  rq_init_comm_if_connected(9, "1")
  rq_init_comm_if_connected(2, "2")
  rq_init_comm_if_connected(3, "3")
  rq_init_comm_if_connected(4, "4")
  rq_print_connected_grippers()
  rq_gripper_communication_thread = run rq_gripper_communication()
  set_closed_norm(97.6470588235294, "1")
  set_open_norm(1.1764705882352942, "1")
  set_closed_mm(0.0, "1")
  set_open_mm(53.0, "1")
  set_closed_norm(100.0, "2")
  set_open_norm(0.0, "2")
  set_closed_mm(0.0, "2")
  set_open_mm(50.0, "2")
  set_closed_norm(100.0, "3")
  set_open_norm(0.0, "3")
  set_closed_mm(0.0, "3")
  set_open_mm(50.0, "3")
  set_closed_norm(100.0, "4")
  set_open_norm(0.0, "4")
  set_closed_mm(0.0, "4")
  set_open_mm(50.0, "4")
  rq_current_limit_enabled = False
  while(not rq_gripper_communication_thread_started):
      sleep(0.008)
  end
  # end: URCap Installation Node
  step_count_652fcfe5_f3e5_4323_a28e_c4dd7c99f65c = 0.0
  thread Step_Counter_Thread_2d5c0d0e_2884_4a5b_ab92_48b0595c18f1():
    while (True):
      step_count_652fcfe5_f3e5_4323_a28e_c4dd7c99f65c = step_count_652fcfe5_f3e5_4323_a28e_c4dd7c99f65c + 1.0
      sync()
    end
  end
  run Step_Counter_Thread_2d5c0d0e_2884_4a5b_ab92_48b0595c18f1()
  global DEV_CEN_PosRtr=0
  $ 2 "BeforeStart"
  $ 3 "Centrifuge≔rpc_factory('xmlrpc','http://192.168.12.125:50002')"
  global Centrifuge=rpc_factory("xmlrpc","http://192.168.12.125:50002")
  $ 4 "Action≔'What to do?'"
  global Action=request_integer_from_primary_client("What to do?")
  $ 5 "Robot Program"
  $ 6 "Handling"
  $ 44 "'===================='"
  # '===================='
  $ 45 "Switch Action"
  switch_1 = Action
  $ 46 "Case 5"
  if (5 == switch_1):
    $ 47 "Open"
    $ 48 "Centrifuge.open_hatch()"
    Centrifuge.open_hatch()
  elif (6 == switch_1):
    $ 49 "Case 6"
    $ 50 "Close"
    $ 51 "Centrifuge.close_hatch()"
    Centrifuge.close_hatch()
  elif (7 == switch_1):
    $ 52 "Case 7"
    $ 53 "Load"
    $ 54 "DEV_CEN_CmdRslt≔Centrifuge.move_rotor(DEV_CEN_PosRtr)"
    global DEV_CEN_CmdRslt=Centrifuge.move_rotor(DEV_CEN_PosRtr)
    $ 55 "If JNT_S≠[0,0,0,0,0,0]"
    if (JNT_S != [0,0,0,0,0,0]):
      $ 56 "MoveJ"
      $ 57 "JNT_S" "breakAfter"
      movej(JNT_S, a=1.3962634015954636, v=1.5707963267948966, r=0.05)
    end
    $ 58 "MoveJ"
    $ 59 "If PSE_A_H≠p[0,0,0,0,0,0]"
    if (PSE_A_H != p[0,0,0,0,0,0]):
      $ 60 "PSE_A_H" "breakAfter"
      movej(pose_trans(FRM_Reference, PSE_A_H), a=1.3962634015954636, v=1.5707963267948966, r=0.02)
    end
    $ 61 "PSE_A" "breakAfter"
    movej(pose_trans(FRM_Reference, PSE_A), a=1.3962634015954636, v=1.5707963267948966)
    $ 62 "If Centrifuge.posreached(DEV_CEN_PosRtr)"
    if (Centrifuge.posreached(DEV_CEN_PosRtr)):
      $ 63 "MoveL"
      $ 64 "If PSE_T_H≠p[0,0,0,0,0,0]"
      if (PSE_T_H != p[0,0,0,0,0,0]):
        $ 65 "PSE_T_H" "breakAfter"
        movel(pose_trans(FRM_Reference, PSE_T_H), a=1.2, v=0.3)
      end
      $ 66 "PSE_T" "breakAfter"
      global move_thread_flag_66=0
      thread move_thread_66():
        enter_critical
        move_thread_flag_66 = 1
        movel(pose_trans(FRM_Reference, PSE_T), a=1.2, v=0.075)
        move_thread_flag_66 = 2
        exit_critical
      end
      move_thread_flag_66 = 0
      move_thread_han_66 = run move_thread_66()
      while (True):
        local targetTcpDirection=get_target_tcp_speed()
        local stepsToRetract=tool_contact(direction=targetTcpDirection)
        if (stepsToRetract > 0):
          kill move_thread_han_66
          stopl(0.5)
          local backTrackMovement=get_actual_joint_positions_history(stepsToRetract)
          local contactPose=get_forward_kin(backTrackMovement)
          local posDir=[targetTcpDirection[0],targetTcpDirection[1],targetTcpDirection[2]]
          local retractTo=contactPose
          if (norm(posDir) > 1e-6):
            local normalizedPosDir=normalize(posDir)
            local additionalRetraction=p[normalizedPosDir[0] * 0.001, normalizedPosDir[1] * 0.001, normalizedPosDir[2] * 0.001, 0, 0, 0]
            retractTo = pose_sub(contactPose, additionalRetraction)
          end
          movel(retractTo, a=0.5, v=0.1)
          $ 67 "Until (tool_contact_detection)"
          $ 68 "EOAT"
          # begin: URCap Program Node
          #   Source: Robotiq_Grippers, 3.11.2.92906, Robotiq Inc.
          #   Type: Gripper
          $ 69 "Gripper Move5mm (1)"
          if not(gripper_connected[0]):
            popup("Gripper 1 must be connected to run this program.", "No connection", False, True, True)
          end
          if not(rq_is_gripper_activated("1")):
            popup("Gripper 1 is not activated. Go to Installation tab > Gripper to activate it and run the program again.", "Not activated", False, True, True)
          end
          rq_set_pos_spd_for(226, 128, 64, "1")
          rq_wait_pos_spe_for_request(226, 128, 64, "1")
          rq_go_to("1")
          rq_wait("1")
          # end: URCap Program Node
          $ 70 "Force"
          sleep(0.02)
          zero_ftsensor()
          force_mode(tool_pose(), [0, 0, 0, 0, 0, 1], [0.0, 0.0, 0.0, 0.0, 0.0, 0.0], 2, [0.1, 0.1, 0.1, 0.3490658503988659, 0.3490658503988659, 3.141592653589793])
          $ 71 "PSE_T" "noBreak"
          movel(pose_trans(FRM_Reference, PSE_T), a=1.2, v=0.01)
          end_force_mode()
          stopl(5.0)
          break
        end
        sleep(1.0E-10)
        if (move_thread_flag_66 > 1):
          join move_thread_han_66
          break
        end
        sync()
      end
      $ 72 "EOAT"
      # begin: URCap Program Node
      #   Source: Robotiq_Grippers, 3.11.2.92906, Robotiq Inc.
      #   Type: Gripper
      $ 73 "Gripper Move15mm (1)"
      if not(gripper_connected[0]):
        popup("Gripper 1 must be connected to run this program.", "No connection", False, True, True)
      end
      if not(rq_is_gripper_activated("1")):
        popup("Gripper 1 is not activated. Go to Installation tab > Gripper to activate it and run the program again.", "Not activated", False, True, True)
      end
      rq_set_pos_spd_for(179, 128, 128, "1")
      rq_wait_pos_spe_for_request(179, 128, 128, "1")
      rq_go_to("1")
      rq_wait("1")
      # end: URCap Program Node
      $ 74 "If PSE_R_H≠p[0,0,0,0,0,0]"
      if (PSE_R_H != p[0,0,0,0,0,0]):
        $ 75 "PSE_R" "breakAfter"
        movel(pose_trans(FRM_Reference, PSE_R), a=1.2, v=0.3, r=0.01)
        $ 76 "PSE_R_H" "breakAfter"
        movel(pose_trans(FRM_Reference, PSE_R_H), a=1.2, v=0.3)
      else:
        $ 77 "Else" "noBreak"
        $ 78 "PSE_R" "breakAfter"
        movel(pose_trans(FRM_Reference, PSE_R), a=1.2, v=0.3)
      end
    end
  elif (8 == switch_1):
    $ 79 "Case 8"
    $ 80 "Unload"
    $ 81 "DEV_CEN_CmdRslt≔Centrifuge.move_rotor(DEV_CEN_PosRtr)"
    global DEV_CEN_CmdRslt=Centrifuge.move_rotor(DEV_CEN_PosRtr)
    $ 82 "If JNT_S≠[0,0,0,0,0,0]"
    if (JNT_S != [0,0,0,0,0,0]):
      $ 83 "MoveJ"
      $ 84 "JNT_S" "breakAfter"
      movej(JNT_S, a=1.3962634015954636, v=1.5707963267948966, r=0.05)
    end
    $ 85 "MoveJ"
    $ 86 "If PSE_A_H≠p[0,0,0,0,0,0]"
    if (PSE_A_H != p[0,0,0,0,0,0]):
      $ 87 "PSE_A_H" "breakAfter"
      movej(pose_trans(FRM_Reference, PSE_A_H), a=1.3962634015954636, v=1.5707963267948966, r=0.02)
    end
    $ 88 "PSE_A" "breakAfter"
    movej(pose_trans(FRM_Reference, PSE_A), a=1.3962634015954636, v=1.5707963267948966)
    $ 89 "EOAT"
    # begin: URCap Program Node
    #   Source: Robotiq_Grippers, 3.11.2.92906, Robotiq Inc.
    #   Type: Gripper
    $ 90 "Gripper Move15mm (1)"
    if not(gripper_connected[0]):
      popup("Gripper 1 must be connected to run this program.", "No connection", False, True, True)
    end
    if not(rq_is_gripper_activated("1")):
      popup("Gripper 1 is not activated. Go to Installation tab > Gripper to activate it and run the program again.", "Not activated", False, True, True)
    end
    rq_set_pos_spd_for(179, 128, 128, "1")
    rq_wait_pos_spe_for_request(179, 128, 128, "1")
    rq_go_to("1")
    rq_wait("1")
    # end: URCap Program Node
    $ 91 "If Centrifuge.posreached(DEV_CEN_PosRtr)"
    if (Centrifuge.posreached(DEV_CEN_PosRtr)):
      $ 92 "MoveL"
      $ 93 "PSE_T" "breakAfter"
      movel(pose_trans(FRM_Reference, PSE_T), a=1.2, v=0.1)
      $ 94 "EOAT"
      # begin: URCap Program Node
      #   Source: Robotiq_Grippers, 3.11.2.92906, Robotiq Inc.
      #   Type: Gripper
      $ 95 "Gripper Close (1)"
      if not(gripper_connected[0]):
        popup("Gripper 1 must be connected to run this program.", "No connection", False, True, True)
      end
      if not(rq_is_gripper_activated("1")):
        popup("Gripper 1 is not activated. Go to Installation tab > Gripper to activate it and run the program again.", "Not activated", False, True, True)
      end
      rq_set_pos_spd_for(255, 128, 128, "1")
      rq_wait_pos_spe_for_request(255, 128, 128, "1")
      rq_go_to("1")
      rq_wait("1")
      # end: URCap Program Node
      $ 96 "If PSE_R_H≠p[0,0,0,0,0,0]"
      if (PSE_R_H != p[0,0,0,0,0,0]):
        $ 97 "PSE_R" "breakAfter"
        movel(pose_trans(FRM_Reference, PSE_R), a=1.2, v=0.3, r=0.01)
        $ 98 "PSE_R_H" "breakAfter"
        movel(pose_trans(FRM_Reference, PSE_R_H), a=1.2, v=0.3)
      else:
        $ 99 "Else" "noBreak"
        $ 100 "PSE_R" "breakAfter"
        movel(pose_trans(FRM_Reference, PSE_R), a=1.2, v=0.3)
      end
    end
  elif (9 == switch_1):
    $ 101 "Case 9"
    $ 102 "Start"
    $ 103 "Centrifuge.start()"
    Centrifuge.start()
  elif (10 == switch_1):
    $ 104 "Case 10"
    $ 105 "Stop"
    $ 106 "Centrifuge.stop()"
    Centrifuge.stop()
  end
  $ 107 "'===================='"
  # '===================='
  $ 108 "PostSettings"
  $ 109 "OBJ_Picked≔rq_is_object_detected()"
  global OBJ_Picked= rq_is_object_detected ()
  $ 110 "Action≔0"
  global Action=0
  $ 111 "Action_Info≔''"
  global Action_Info=""
end
